RoboDK station: Lab02_mariposa_polar.rdk

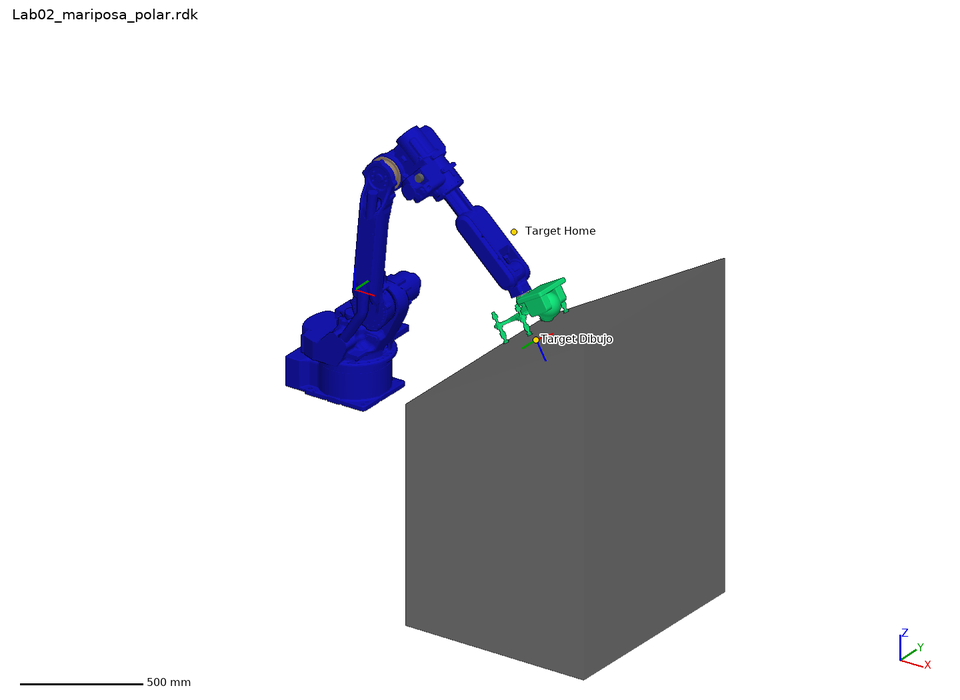
[picture v0: the station drawn from its stored meshes, robots at their saved joint values, targets as dots, program paths as lines]
Station Robodk (2) (saved by RoboDK 6.1.1). Poses are relative to the parent item; angles as X-Y-Z fixed-axis rotations.
  - frame Motoman MH6 Base at (0, 0, 450) mm
    - robot Motoman MH6: 6 axes, payload 6 kg, reach 1422 mm, repeatability 0.08 mm, weight 130 kg
        modified DH rows (alpha deg, a mm, theta deg, d mm): 0, 0, 0, 450; -90, 152, -90, 0; 0, 614, 0, 0; -90, 155, 0, 640; 90, 0, 90, 0; -90, 0, 0, 95
        base shift (0, 0, -450) mm
        joint limits [-170, -90, -175, -180, -45, -360] to [170, 155, 250, 180, 225, 360]; home [0, 0, 0, 0, 0, 0]; saved at [0.229, 5.197, -37.914, 0.394, 73.111, -0.575]
      - tool Ventosas, TCP at (0, 0, 190) mm, size 250 x 290 x 148 mm
    - target   Target Home (joint target) at (792, 0, 484) mm, rotated rx -180 ry 0 rz 0 deg; joints [0, 0, 0, 0, 0, 0] of Motoman MH6
    - target Target Dibujo (Cartesian target) at (900, 0, 25) mm, rotated rx 180 ry 0 rz 0 deg; joints [0, 14.531, -24.666, 0, 39.198, 0] of Motoman MH6
  - object CAJA2 at (1600, 500, 300) mm, rotated rx 180 ry 0 rz 0 deg, size 886.4 x 1000 x 1511.7 mm, geometry from CAJA2.stp
  - Python program RosPolar (listed below)
  - frame Frame_from_Target1 at (900, 0, 477) mm, rotated rx 180 ry -30 rz 0 deg

--- Python program RosPolar ---
## =====================================================================
#  Laboratorio No. 02 - Robótica Industrial 2026-II - UNAL
#  Trayectoria polar en RoboDK + Motoman MH6 (controlador DX100)
#  Figura: MARIPOSA POLAR (curva de Temple Fay)
#           r(t) = e^(sin t) − 2·cos(4t) + sin^5((2t − π)/24),  t ∈ [0, 12π]
#  Integrantes: Alexandra Garavito y David Ruiz
# =====================================================================
from robodk.robolink import *    # API para comunicarse con RoboDK
from robodk.robomath import *    # transl(), rotx(), etc.
import math
import numpy as np

# ---------------------------------------------------------------------
# 0) MODO DE EJECUCIÓN
#    False -> SIMULACIÓN: se usa la herramienta virtual y NO se conecta
#             al robot real (equivale a comentar el bloque de conexión).
#    True  -> ROBOT REAL: se conecta al DX100 y NO se fuerza la herramienta
#             virtual (equivale a comentar setPoseTool).
# ---------------------------------------------------------------------
MODO_REAL = False
VERIFICAR_ALCANCE = True   # Antes de mover, comprueba que TODOS los puntos sean alcanzables

NOMBRE_FRAME = "Frame_from_Target1"   # Frame con origen SOBRE el papel (centro del dibujo)
NOMBRE_HERRAMIENTA = "Ventosas"       # Herramienta virtual de la estación (solo simulación)
NOMBRE_HOME = "Target Home"           # Target creado PRIMERO en la estación (nombre exacto del árbol)

# ---------------------------------------------------------------------
# 1) PARÁMETROS DE LA FIGURA
# ---------------------------------------------------------------------
A = 150.0              # Radio máximo [mm]: r = A * r_raw / max|r_raw|  (max|r_raw| ≈ 5.05)
                       # -> figura ≈ 217 x 191 mm (x: ±108, y: -74 a 117)
T_FINAL = 12 * math.pi # 6 vueltas para que aparezcan las alas "dobles"
NUM_PUNTOS = 1000      # Longitud total ≈ 6448 mm -> segmentos ≈ 6.4 mm.
                       # Balance red/forma: con 2000 pts (3.2 mm) se duplican los paquetes por
                       # Ethernet y el robot hace "pare-arranque"; con ~400 (16 mm) los lóbulos
                       # pequeños del centro se ven poligonales.

# Alturas: SIEMPRE distancias positivas (buena práctica). El signo lo pone pose().
Z_SEGURA = 50.0        # Altura de aproximación / salida [mm]
Z_LEVANTE = 10.0       # Levante corto entre letras [mm]

# Velocidades
V_LINEAL_APROX = 150.0   # mm/s  (aproximación, subir/bajar)
V_JOINT = 30.0           # deg/s (MoveJ: Home y aproximación)
V_DIBUJO = 60.0          # mm/s  (trazo). Con segmentos de 6.4 mm -> ~107 ms por punto,
                         # tiempo suficiente para que cada paquete llegue al DX100.
                         # Trazo de la mariposa ≈ 6448/60 ≈ 1 min 50 s.

# Redondeo (zona de aproximación). En el DX100 se traduce a nivel de posicionamiento PL.
REDONDEO_DIBUJO = 1.0    # mm. Debe ser MENOR que la mitad del segmento (6.4/2 ≈ 3.2 mm).
                         # Con 5 mm (código original) la zona era más grande que los
                         # segmentos y la figura se deformaba.
REDONDEO_PRECISO = -1    # -1 = sin redondeo (llega exacto al punto). Para Home, bajar y subir.

# Nombres con TextPath (matplotlib) debajo de la mariposa (opcional)
ESCRIBIR_TEXTO = True
LINEAS_TEXTO = ["ALEXANDRA", "DAVID"]   # Integrantes del grupo (una línea por nombre)
ALTURA_TEXTO = 16.0      # mm (en una sola línea las letras quedarían de ~10 mm)
ANCHO_MAX_TEXTO = 170.0  # mm
Y_TEXTO = -90.0          # mm (borde superior de la 1.ª línea; la mariposa llega hasta y ≈ -74 mm)
INTERLINEADO = 6.0       # mm entre líneas

# ---------------------------------------------------------------------
# 2) GEOMETRÍA (Python puro, se puede probar sin RoboDK)
# ---------------------------------------------------------------------
# El frame se creó desde un target ("Frame_from_Target1"), por lo tanto su eje Z
# es el Z de la herramienta y apunta HACIA el papel. "Subir" es ir en -Z.
# (Si su frame tuviera Z hacia arriba, cambie a +1 y agregue rotx(pi) en pose()).
SIGNO_SUBIR = -1

# Giro del dibujo (mariposa + nombres) dentro del plano de la cara, en grados.
# Positivo = antihorario visto de frente a la cara. 180 = voltear de cabeza.
ROTACION_DIBUJO = -90.0


def pose(x, y, altura=0.0):
    """Pose en el frame de trabajo. altura = distancia (positiva) sobre el papel.
    Si el eje Z del frame apunta HACIA el papel, al mirar desde arriba el plano XY
    queda en espejo; se invierte Y para que la mariposa y los nombres se lean bien."""
    if ROTACION_DIBUJO:
        c = math.cos(math.radians(ROTACION_DIBUJO))
        s_ = math.sin(math.radians(ROTACION_DIBUJO))
        x, y = c * x - s_ * y, s_ * x + c * y
    if SIGNO_SUBIR == -1:
        y = -y
    return transl(x, y, SIGNO_SUBIR * altura)


def puntos_mariposa(A, n_puntos, t_final=T_FINAL, muestras=200000):
    """Mariposa polar normalizada (mismo cálculo que en GeoGebra/RosPolar.py).
    Devuelve n_puntos+1 puntos (x, y) [mm] separados la MISMA distancia sobre
    la curva (remuestreo por longitud de arco). Con linspace en t los segmentos
    van de <1 mm a >15 mm; así todos miden igual y un único redondeo sirve."""
    # a) Muestreo denso en t
    t_values = np.linspace(0, t_final, muestras + 1)
    r_raw = (np.exp(np.sin(t_values))
             - 2 * np.cos(4 * t_values)
             + np.sin((2 * t_values - math.pi) / 24) ** 5)
    r = A * r_raw / np.max(np.abs(r_raw))          # normalización del radio
    x = r * np.cos(t_values)
    y = r * np.sin(t_values)
    # b) Longitud de arco acumulada
    s = np.concatenate(([0.0], np.cumsum(np.hypot(np.diff(x), np.diff(y)))))
    total = s[-1]
    # c) n_puntos segmentos de igual longitud
    s_obj = np.linspace(0, total, n_puntos + 1)
    xs = np.interp(s_obj, s, x)
    ys = np.interp(s_obj, s, y)
    return list(zip(xs.tolist(), ys.tolist())), total


def contornos_texto(texto, altura, ancho_max, y_superior, sep_min=0.8):
    """Contornos de las letras con matplotlib.textpath.TextPath, en mm,
    centrados en x = 0 y con el borde superior en y_superior."""
    from matplotlib.textpath import TextPath
    from matplotlib.font_manager import FontProperties
    tp = TextPath((0, 0), texto, size=1.0, prop=FontProperties(family="DejaVu Sans", weight="bold"))
    polys = [p for p in tp.to_polygons() if len(p) > 1]
    xs = [p[0] for poly in polys for p in poly]
    ys = [p[1] for poly in polys for p in poly]
    xmin, xmax, ymin, ymax = min(xs), max(xs), min(ys), max(ys)
    esc = min(altura / (ymax - ymin), ancho_max / (xmax - xmin))
    xc = (xmin + xmax) / 2.0
    contornos = []
    for poly in polys:
        pts = [((px - xc) * esc, (py - ymax) * esc + y_superior) for px, py in poly]
        # Quitar puntos casi repetidos (no saturar la red con segmentos < sep_min)
        limpio = [pts[0]]
        for p in pts[1:]:
            if math.hypot(p[0] - limpio[-1][0], p[1] - limpio[-1][1]) >= sep_min:
                limpio.append(p)
        if limpio[-1] != pts[0]:
            limpio.append(pts[0])          # cerrar el contorno
        contornos.append(limpio)
    return contornos


# ---------------------------------------------------------------------
# 3) PROGRAMA PRINCIPAL (RoboDK)
# ---------------------------------------------------------------------
def main():
    RDK = Robolink()

    robot = RDK.ItemUserPick("Selecciona un robot", ITEM_TYPE_ROBOT)
    if not robot.Valid():
        raise Exception("No se ha seleccionado un robot válido.")

    if MODO_REAL:
        # ---------- CONEXIÓN AL ROBOT REAL (comentar en simulación) ----------
        if robot.Connect() != 1:          # Connect() devuelve 1 si conectó
            raise Exception("No se pudo conectar. Verifique modo REMOTE, IP y servos.")
        estado, msg = robot.ConnectedState()   # devuelve (código, mensaje)
        if estado != ROBOTCOM_READY:
            raise Exception("El robot no está listo: " + msg)
        RDK.setRunMode(RUNMODE_RUN_ROBOT)
        print("Robot real conectado:", msg)
    else:
        # ---------- HERRAMIENTA VIRTUAL (comentar en real) ----------
        RDK.setRunMode(RUNMODE_SIMULATE)
        herramienta = RDK.Item(NOMBRE_HERRAMIENTA, ITEM_TYPE_TOOL)
        if not herramienta.Valid():
            herramienta = robot.getLink(ITEM_TYPE_TOOL)   # herramienta activa
        robot.setPoseTool(herramienta)
        print("Modo simulación con herramienta:", herramienta.Name())

    frame = RDK.Item(NOMBRE_FRAME, ITEM_TYPE_FRAME)
    if not frame.Valid():
        raise Exception(f'No se encontró el Frame "{NOMBRE_FRAME}" en la estación.')
    robot.setPoseFrame(frame)

    # Target Home: se crea PRIMERO en RoboDK (Ctrl+T) y aquí solo se llama por su nombre
    home = RDK.Item(NOMBRE_HOME, ITEM_TYPE_TARGET)
    if not home.Valid():
        raise Exception(f'No se encontró el target "{NOMBRE_HOME}". Créelo en la estación antes de ejecutar.')

    # ---------- Puntos de toda la rutina (se calculan ANTES de mover) ----------
    mariposa, perimetro = puntos_mariposa(A, NUM_PUNTOS)
    contornos = []
    if ESCRIBIR_TEXTO:
        try:
            for i, linea in enumerate(LINEAS_TEXTO):
                y_sup = Y_TEXTO - i * (ALTURA_TEXTO + INTERLINEADO)
                contornos += contornos_texto(linea, ALTURA_TEXTO, ANCHO_MAX_TEXTO, y_sup)
        except ImportError:
            print("matplotlib no está instalado en el Python de RoboDK: se omite el texto.")

    todos = mariposa + [p for c in contornos for p in c]
    xs = [p[0] for p in todos]
    ys = [p[1] for p in todos]
    print(f"Mariposa: {NUM_PUNTOS} segmentos de {perimetro / NUM_PUNTOS:.2f} mm")
    print(f"Rotación del dibujo: {ROTACION_DIBUJO:.0f}°")
    print(f"Área que ocupa el dibujo en el frame: x [{min(xs):.0f}, {max(xs):.0f}] mm,"
          f" y [{min(ys):.0f}, {max(ys):.0f}] mm")

    # ---------- Verificación de alcance (no mueve el robot) ----------
    if VERIFICAR_ALCANCE:
        herr_pose = robot.PoseTool()
        ref_pose = robot.PoseFrame()
        q_prev = home.Joints().list()
        revisar = [(todos[0][0], todos[0][1], Z_SEGURA)]           # aproximación
        revisar += [(x, y, 0.0) for (x, y) in todos]                # puntos sobre el papel
        revisar += [(todos[-1][0], todos[-1][1], Z_SEGURA)]         # salida
        for (x, y, h) in revisar:
            q = robot.SolveIK(pose(x, y, h), q_prev, herr_pose, ref_pose).list()
            if len(q) < 6:
                raise Exception(f"Punto NO alcanzable: x={x:.1f}, y={y:.1f}, altura={h:.0f} mm. "
                                "Acerque el frame al robot o reduzca A.")
            q_prev = q[:6]
        print("Verificación OK: todos los puntos son alcanzables.")

    def ir_a_home():
        robot.setRounding(REDONDEO_PRECISO)      # llegar exacto a Home (sin redondeo)
        robot.setSpeed(V_LINEAL_APROX, V_JOINT)
        robot.MoveJ(home.Joints())   # articulaciones guardadas en el target (evita TargetReachError)

    def trazar(puntos, altura_entrada, altura_salida):
        """Aproxima, baja, recorre la polilínea con redondeo y sube."""
        x0, y0 = puntos[0]
        robot.setRounding(REDONDEO_PRECISO)
        robot.setSpeed(V_LINEAL_APROX, V_JOINT)
        robot.MoveL(pose(x0, y0, altura_entrada))   # encima del primer punto
        robot.MoveL(pose(x0, y0, 0.0))              # bajar al papel
        robot.setSpeed(V_DIBUJO)
        robot.setRounding(REDONDEO_DIBUJO)
        for (x, y) in puntos[1:]:
            robot.MoveL(pose(x, y, 0.0))
        robot.setRounding(REDONDEO_PRECISO)
        robot.setSpeed(V_LINEAL_APROX)
        xf, yf = puntos[-1]
        robot.MoveL(pose(xf, yf, altura_salida))    # subir

    # ---------------- RUTINA: Home -> mariposa -> nombres -> Home ----------------
    ir_a_home()                            # 1) INICIO en Home

    x0, y0 = mariposa[0]
    robot.MoveJ(pose(x0, y0, Z_SEGURA))    # 2) aproximación sobre el PRIMER punto (no el centro)
    trazar(mariposa, Z_SEGURA, Z_SEGURA)   # 3) mariposa (for con redondeo pequeño)

    for k, c in enumerate(contornos):      # 4) nombres, letra por letra
        salida = Z_SEGURA if k == len(contornos) - 1 else Z_LEVANTE
        trazar(c, Z_LEVANTE, salida)

    ir_a_home()                            # 5) FIN en Home
    print(f"¡Mariposa polar completada en el frame '{NOMBRE_FRAME}'!")


if __name__ == "__main__":
    main()
